TYPE "ST_AirPressureParCfg"
VERSION : 0.1
   STRUCT
      SchemaVersion : UInt := 1;
      ConflictTime : Time := T#500MS;
   END_STRUCT;

END_TYPE

